(* IEC 61131-3 sources: NachHouse_TST/API/pilot_Api_V11 (part 2) *)

(* ---- 03_Nh_Api_ENGINE.st ---- *)
// Single-owner transaction engine, snapshots, diffs and room operations.
// SK: Transakcny automat jedneho vlastnika, snapshoty, diffy a room operacie.

FUNCTION NhApiClearRoom : BOOL
   // Clears configuration and state of one internal room slot. SK: Vynuluje konfiguraciu a stav jedneho interneho room slotu.
   VAR_INPUT
      Index : UINT; // Internal model-device slot 1..800. SK: Interny slot modeloveho zariadenia 1..800.
   END_VAR
   NhRoomsConfig[Index].Used := FALSE;
   NhRoomsConfig[Index].RoomId := 0;
   NhRoomsConfig[Index].Name := '';
   NhRoomsConfig[Index].ProjectName := '';
   NhRoomsConfig[Index].IconId := 0;
   NhRoomsConfig[Index].SortDefault := 0;
   NhRoomsState[Index].RoomId := 0;
   NhRoomsState[Index].Temperature := 0.0;
   NhRoomsState[Index].Humidity := 0.0;
   NhRoomsState[Index].Presence := FALSE;
   NhRoomsState[Index].DayPhase := 140;
   NhRoomsState[Index].CategoryMask := 0;
   NhRoomsState[Index].AlarmLevel := 0;
   NhRoomsState[Index].Online := FALSE;
   NhRoomsState[Index].Twilight := FALSE;
   NhApiClearRoom := TRUE;
END_FUNCTION

FUNCTION NhApiInitialize : BOOL
   // Initializes API buffers, handshake and deterministic pilot data once. SK: Jednorazovo inicializuje API buffery, handshake a deterministicke pilotne data.
   VAR
      Index : UINT; // Initialization index. SK: Inicializacny index.
   END_VAR
   NhApiInitialize := NhApiInitialized;
   IF NhApiInitialized THEN RETURN; END_IF;

   NhApiClearBuffer(Buffer := ADR(NhApiTX), Length := NH_API_TX_BYTE_CAPACITY);
   NhApiClearBuffer(Buffer := ADR(NhApiRX), Length := NH_API_RX_BYTE_CAPACITY);
   FOR Index := 1 TO NH_API_MAX_ROOMS DO
      NhApiClearRoom(Index := Index);
   END_FOR;

   FOR Index := 1 TO 30 DO
      NhRoomsConfig[Index].Used := TRUE;
      NhRoomsConfig[Index].RoomId := UINT_TO_UDINT(Index);
      NhRoomsConfig[Index].ProjectName := 'TEST';
      NhRoomsConfig[Index].IconId := SEL(Index >= 26, 16, 19);
      NhRoomsConfig[Index].SortDefault := Index;
      CASE Index OF
         1: NhRoomsConfig[Index].Name := 'Hall 1'; NhRoomsConfig[Index].ProjectName := '1.08';
         2: NhRoomsConfig[Index].Name := 'Kitchen'; NhRoomsConfig[Index].ProjectName := '1.07';
         3: NhRoomsConfig[Index].Name := 'Corridor 1'; NhRoomsConfig[Index].ProjectName := '1.04';
         4: NhRoomsConfig[Index].Name := 'Bathroom 1'; NhRoomsConfig[Index].ProjectName := '1.06';
         5: NhRoomsConfig[Index].Name := 'WC'; NhRoomsConfig[Index].ProjectName := '1.05';
         6: NhRoomsConfig[Index].Name := 'Bedroom'; NhRoomsConfig[Index].ProjectName := '1.09';
         7: NhRoomsConfig[Index].Name := 'Boiler'; NhRoomsConfig[Index].ProjectName := '1.03';
         8: NhRoomsConfig[Index].Name := 'Living room'; NhRoomsConfig[Index].ProjectName := '1.01';
         9: NhRoomsConfig[Index].Name := 'Corridor 1F'; NhRoomsConfig[Index].ProjectName := '1.02';
         10: NhRoomsConfig[Index].Name := 'Room 2.07'; NhRoomsConfig[Index].ProjectName := '2.07';
         11: NhRoomsConfig[Index].Name := 'Kitchen 2F'; NhRoomsConfig[Index].ProjectName := '2.03';
         12: NhRoomsConfig[Index].Name := 'Room 2.06'; NhRoomsConfig[Index].ProjectName := '2.06';
         13: NhRoomsConfig[Index].Name := 'Bathroom 2F'; NhRoomsConfig[Index].ProjectName := '2.05';
         14: NhRoomsConfig[Index].Name := 'Entrance hall'; NhRoomsConfig[Index].ProjectName := '0.01';
         15: NhRoomsConfig[Index].Name := 'Garage'; NhRoomsConfig[Index].ProjectName := '0.02';
         16: NhRoomsConfig[Index].Name := 'Storage'; NhRoomsConfig[Index].ProjectName := '0.03';
         17: NhRoomsConfig[Index].Name := 'Basement corridor'; NhRoomsConfig[Index].ProjectName := '0.04';
         18: NhRoomsConfig[Index].Name := 'Office'; NhRoomsConfig[Index].ProjectName := '1.10';
         19: NhRoomsConfig[Index].Name := 'Wardrobe'; NhRoomsConfig[Index].ProjectName := '1.11';
         20: NhRoomsConfig[Index].Name := 'Fitness'; NhRoomsConfig[Index].ProjectName := '0.06';
         21: NhRoomsConfig[Index].Name := 'Technical'; NhRoomsConfig[Index].ProjectName := '0.07';
         22: NhRoomsConfig[Index].Name := 'Wine room'; NhRoomsConfig[Index].ProjectName := '0.08';
         23: NhRoomsConfig[Index].Name := 'Guest room'; NhRoomsConfig[Index].ProjectName := '2.01';
         24: NhRoomsConfig[Index].Name := 'Children 1'; NhRoomsConfig[Index].ProjectName := '2.02';
         25: NhRoomsConfig[Index].Name := 'Children 2'; NhRoomsConfig[Index].ProjectName := '2.04';
         26: NhRoomsConfig[Index].Name := 'Terrace'; NhRoomsConfig[Index].ProjectName := 'E.01';
         27: NhRoomsConfig[Index].Name := 'Gazebo'; NhRoomsConfig[Index].ProjectName := 'E.02';
         28: NhRoomsConfig[Index].Name := 'Pool'; NhRoomsConfig[Index].ProjectName := 'E.03';
         29: NhRoomsConfig[Index].Name := 'Garden'; NhRoomsConfig[Index].ProjectName := 'E.04';
         30: NhRoomsConfig[Index].Name := 'Sauna'; NhRoomsConfig[Index].ProjectName := '0.09';
      END_CASE;
      NhRoomsState[Index].RoomId := UINT_TO_UDINT(Index);
      NhRoomsState[Index].Temperature := 20.0 + UINT_TO_REAL(Index) * 0.1;
      NhRoomsState[Index].Humidity := 40.0 + UINT_TO_REAL(Index MOD 15);
      NhRoomsState[Index].Presence := (Index MOD 4) = 0;
      CASE Index MOD 4 OF
         0: NhRoomsState[Index].DayPhase := 140;
         1: NhRoomsState[Index].DayPhase := 142;
         2: NhRoomsState[Index].DayPhase := 144;
         3: NhRoomsState[Index].DayPhase := 146;
      END_CASE;
      NhRoomsState[Index].CategoryMask := UINT_TO_DWORD(Index MOD 8);
      NhRoomsState[Index].AlarmLevel := 0;
      NhRoomsState[Index].Online := (Index MOD 3) <> 0;
      NhRoomsState[Index].Twilight := (Index MOD 3) <> 1;
   END_FOR;

   FOR Index := 1 TO NH_API_MAX_ROOMS DO
      NhConfigShadow[Index] := NhRoomsConfig[Index];
      NhStateShadow[Index] := NhRoomsState[Index];
   END_FOR;

   // Deterministic compact LOAD_800 device model. SK: Deterministicky kompaktny model 800 zariadeni.
   FOR Index := 1 TO NH_LOAD_DEVICE_COUNT DO
      IF Index <= 300 THEN
         NhLoadDevices[Index] := 16#01000064; // light, level 100
      ELSIF Index <= 420 THEN
         NhLoadDevices[Index] := 16#02000064; // roller, position 100
      ELSIF Index <= 520 THEN
         NhLoadDevices[Index] := 16#030000D2; // heating, 21.0 C
      ELSIF Index <= 600 THEN
         NhLoadDevices[Index] := 16#040000DC; // climate, 22.0 C
      ELSIF Index <= 640 THEN
         NhLoadDevices[Index] := 16#05000001; // water, enabled
      ELSE
         NhLoadDevices[Index] := 16#06000000 OR UINT_TO_DWORD(Index MOD 256); // sensor control group
      END_IF;
   END_FOR;

   NhApiInfo.ApiVersion := NH_API_VERSION;
   NhApiInfo.OwnerClientId := 0;
   NhApiInfo.State := NH_API_STATE_IDLE;
   NhActiveOwnerClientId := 0;
   NhExpectedState := NH_API_STATE_IDLE;
   NhTransactionMode := NH_API_MODE_NONE;
   NhTransactionLastMs := NhApiSystemTimeMs();
   NhPublishedFrameId := 0;
   NhCommandResult := NH_API_RESULT_NONE;
   NhResultPending := FALSE;
   NhPendingConfigCount := 0;
   NhPendingStateCount := 0;
   NhSnapshotActive := FALSE;

   NhApiTest.Execute := FALSE;
   NhApiTest.Finished := FALSE;
   NhApiTest.Action := NH_API_TEST_NONE;
   NhApiTest.ResultCode := NH_API_RESULT_NONE;
   NhLoadTest.DepartureActive := FALSE;
   NhLoadTest.LastChangedCount := 0;
   NhLoadTest.LastApplyMs := 0;
   NhLoadTest.Sequence := 0;
   NhApiInitialized := TRUE;
   NhApiInitialize := TRUE;
END_FUNCTION

FUNCTION NhApiBeginFrame : BOOL
   // Clears TX and writes the fixed 40-byte frame header. SK: Vycisti TX a zapise pevnu 40-bajtovu hlavicku ramca.
   VAR_INPUT
      MessageType  : UINT;  // NH_API_MSG_* value. SK: Hodnota NH_API_MSG_*.
      SchemaId     : UINT;  // NH_API_SCHEMA_* value. SK: Hodnota NH_API_SCHEMA_*.
      OwnerClientId: UDINT; // Target owner token; zero is broadcast. SK: Cielovy token vlastnika; nula je broadcast.
      RecordCount  : UINT;  // Number of payload records. SK: Pocet zaznamov payloadu.
      RecordSize   : UINT;  // Fixed size of one payload record. SK: Pevna velkost jedneho payload zaznamu.
      PartIndex    : UINT;  // One-based part index. SK: Index casti cislovany od jedna.
      PartCount    : UINT;  // Total parts in this section. SK: Celkovy pocet casti sekcie.
      ResultCode   : USINT; // NH_API_RESULT_* value. SK: Hodnota NH_API_RESULT_*.
   END_VAR
   VAR
      Buffer      : PTR_TO BYTE; // Byte view of NhApiTX. SK: Bajtovy pohlad na NhApiTX.
      PayloadSize : UDINT;       // Calculated payload size. SK: Vypocitana velkost payloadu.
      TotalSize   : UDINT;       // Header plus payload size. SK: Velkost hlavicky a payloadu.
   END_VAR
   Buffer := ADR(NhApiTX);
   NhApiClearBuffer(Buffer := Buffer, Length := NH_API_TX_BYTE_CAPACITY);
   PayloadSize := UINT_TO_UDINT(RecordCount) * UINT_TO_UDINT(RecordSize);
   TotalSize := UINT_TO_UDINT(NH_API_HEADER_SIZE) + PayloadSize;
   IF TotalSize > UINT_TO_UDINT(NH_API_TX_BYTE_CAPACITY) THEN
      NhApiBeginFrame := FALSE;
      RETURN;
   END_IF;
   NhApiWriteU32(Buffer := Buffer, Offset := 0, Value := DWORD_TO_UDINT(NH_API_MAGIC));
   NhApiWriteU16(Buffer := Buffer, Offset := 4, Value := NH_API_VERSION);
   NhApiWriteU16(Buffer := Buffer, Offset := 6, Value := NH_API_HEADER_SIZE);
   NhApiWriteU16(Buffer := Buffer, Offset := 8, Value := MessageType);
   NhApiWriteU16(Buffer := Buffer, Offset := 10, Value := SchemaId);
   NhApiWriteU32(Buffer := Buffer, Offset := 12, Value := OwnerClientId);
   NhApiWriteU16(Buffer := Buffer, Offset := 16, Value := RecordCount);
   NhApiWriteU16(Buffer := Buffer, Offset := 18, Value := RecordSize);
   NhApiWriteByte(Buffer := Buffer, Offset := 20, Value := WORD_TO_BYTE(UINT_TO_WORD(PartIndex)));
   NhApiWriteByte(Buffer := Buffer, Offset := 21, Value := WORD_TO_BYTE(UINT_TO_WORD(PartCount)));
   NhApiWriteByte(Buffer := Buffer, Offset := 22, Value := USINT_TO_BYTE(ResultCode));
   NhApiWriteByte(Buffer := Buffer, Offset := 23, Value := 0);
   NhApiWriteU32(Buffer := Buffer, Offset := 24, Value := PayloadSize);
   NhApiWriteU32(Buffer := Buffer, Offset := 28, Value := TotalSize);
   NhApiWriteU32(Buffer := Buffer, Offset := 32, Value := 0);
   NhApiWriteU32(Buffer := Buffer, Offset := 36, Value := 0);
   NhApiBeginFrame := TRUE;
END_FUNCTION

FUNCTION NhApiPublishFrame : BOOL
   // Adds CRC and publishes TX by changing State only after the buffer is stable. SK: Doplni CRC a publikuje TX zmenou State az po ustaleni buffera.
   VAR_INPUT
      NextState : UINT; // New persistent handshake step. SK: Novy trvaly handshake krok.
   END_VAR
   VAR
      Buffer    : PTR_TO BYTE; // Byte view of NhApiTX. SK: Bajtovy pohlad na NhApiTX.
      TotalSize : UINT;        // Valid frame byte count. SK: Pocet platnych bajtov ramca.
      Crc       : DWORD;       // CRC32 of the frame. SK: CRC32 ramca.
   END_VAR
   Buffer := ADR(NhApiTX);
   TotalSize := UDINT_TO_UINT(NhApiReadU32(Buffer := Buffer, Offset := 28));
   NhPublishedFrameId := NhPublishedFrameId + 1;
   IF NhPublishedFrameId = 0 THEN NhPublishedFrameId := 1; END_IF;
   NhApiWriteU32(Buffer := Buffer, Offset := 32, Value := NhPublishedFrameId);
   Crc := NhApiFrameCrc32(Buffer := Buffer, Length := TotalSize);
   NhApiWriteU32(Buffer := Buffer, Offset := 36, Value := DWORD_TO_UDINT(Crc));
   NhExpectedState := NextState;
   NhTransactionLastMs := NhApiSystemTimeMs();
   NhApiInfo.State := NextState;
   NhApiPublishFrame := TRUE;
END_FUNCTION

FUNCTION NhApiResetTransaction : BOOL
   // Releases the global mailbox and clears internal sequence state. SK: Uvolni globalny mailbox a vycisti interny stav sekvencie.
   NhApiInfo.OwnerClientId := 0;
   NhApiInfo.State := NH_API_STATE_IDLE;
   NhActiveOwnerClientId := 0;
   NhExpectedState := NH_API_STATE_IDLE;
   NhTransactionMode := NH_API_MODE_NONE;
   NhTransactionLastMs := NhApiSystemTimeMs();
   NhCommandResult := NH_API_RESULT_NONE;
   NhResultPending := FALSE;
   NhPendingConfigCount := 0;
   NhPendingStateCount := 0;
   NhSnapshotActive := FALSE;
   NhApiResetTransaction := TRUE;
END_FUNCTION

FUNCTION NhApiApplyAdd : USINT
   // Adds a room to the first free internal slot. SK: Prida miestnost do prveho volneho interneho slotu.
   VAR_INPUT
      Record : NH_ROOM_CONFIG; // New room configuration. SK: Konfiguracia novej miestnosti.
   END_VAR
   VAR
      Slot : UINT; // Free internal room slot. SK: Volny interny room slot.
   END_VAR
   IF (Record.RoomId = 0) OR (LEN(Record.Name) = 0) THEN NhApiApplyAdd := NH_API_RESULT_INVALID; RETURN; END_IF;
   IF NhApiFindRoom(RoomId := Record.RoomId) <> 0 THEN NhApiApplyAdd := NH_API_RESULT_ALREADY_EXISTS; RETURN; END_IF;
   Slot := NhApiFindFreeRoom();
   IF Slot = 0 THEN NhApiApplyAdd := NH_API_RESULT_NO_FREE_SLOT; RETURN; END_IF;
   NhRoomsConfig[Slot] := Record;
   NhRoomsConfig[Slot].Used := TRUE;
   IF NhRoomsConfig[Slot].IconId = 0 THEN NhRoomsConfig[Slot].IconId := 16; END_IF;
   IF NhRoomsConfig[Slot].SortDefault = 0 THEN NhRoomsConfig[Slot].SortDefault := Slot; END_IF;
   NhRoomsState[Slot].RoomId := Record.RoomId;
   NhRoomsState[Slot].Temperature := 20.0;
   NhRoomsState[Slot].Humidity := 40.0;
   NhRoomsState[Slot].Presence := FALSE;
   NhRoomsState[Slot].DayPhase := 140;
   NhRoomsState[Slot].CategoryMask := 0;
   NhRoomsState[Slot].AlarmLevel := 0;
   NhRoomsState[Slot].Online := TRUE;
   NhRoomsState[Slot].Twilight := FALSE;
   NhApiApplyAdd := NH_API_RESULT_OK;
END_FUNCTION

FUNCTION NhApiApplyDelete : USINT
   // Deletes a room by stable RoomId. SK: Zmaze miestnost podla stabilneho RoomId.
   VAR_INPUT
      RoomId : UDINT; // ID of the room to delete. SK: ID mazanej miestnosti.
   END_VAR
   VAR
      Slot : UINT;   // Located internal slot. SK: Najdeny interny slot.
   END_VAR
   Slot := NhApiFindRoom(RoomId := RoomId);
   IF Slot = 0 THEN NhApiApplyDelete := NH_API_RESULT_NOT_FOUND; RETURN; END_IF;
   NhApiClearRoom(Index := Slot);
   NhApiApplyDelete := NH_API_RESULT_OK;
END_FUNCTION

FUNCTION NhApiApplyConfig : USINT
   // Replaces complete configuration of an existing room. SK: Nahradi celu konfiguraciu existujucej miestnosti.
   VAR_INPUT
      Record : NH_ROOM_CONFIG; // Complete new configuration. SK: Uplna nova konfiguracia.
   END_VAR
   VAR
      Slot : UINT;            // Located internal slot. SK: Najdeny interny slot.
   END_VAR
   Slot := NhApiFindRoom(RoomId := Record.RoomId);
   IF Slot = 0 THEN NhApiApplyConfig := NH_API_RESULT_NOT_FOUND; RETURN; END_IF;
   IF LEN(Record.Name) = 0 THEN NhApiApplyConfig := NH_API_RESULT_INVALID; RETURN; END_IF;
   NhRoomsConfig[Slot] := Record;
   NhRoomsConfig[Slot].Used := TRUE;
   NhApiApplyConfig := NH_API_RESULT_OK;
END_FUNCTION

FUNCTION NhApiApplyState : USINT
   // Replaces complete dynamic state of an existing room. SK: Nahradi cely dynamicky stav existujucej miestnosti.
   VAR_INPUT
      Record : NH_ROOM_STATE; // Complete new state. SK: Uplny novy stav.
   END_VAR
   VAR
      Slot : UINT;           // Located internal slot. SK: Najdeny interny slot.
   END_VAR
   Slot := NhApiFindRoom(RoomId := Record.RoomId);
   IF Slot = 0 THEN NhApiApplyState := NH_API_RESULT_NOT_FOUND; RETURN; END_IF;
   IF (Record.Temperature < -50.0) OR (Record.Temperature > 100.0) OR
      (Record.Humidity < 0.0) OR (Record.Humidity > 100.0) OR (Record.AlarmLevel > 2) THEN
      NhApiApplyState := NH_API_RESULT_INVALID;
      RETURN;
   END_IF;
   NhRoomsState[Slot] := Record;
   NhApiApplyState := NH_API_RESULT_OK;
END_FUNCTION

FUNCTION NhApiApplyCopy : USINT
   // Copies an existing room into a new RoomId. SK: Skopiruje existujucu miestnost do noveho RoomId.
   VAR_INPUT
      SourceRoomId : UDINT;         // Source room ID. SK: ID zdrojovej miestnosti.
      Target       : NH_ROOM_CONFIG;// Target ID and optional replacements. SK: Cielove ID a volitelne nahrady.
   END_VAR
   VAR
      SourceSlot : UINT; // Source internal slot. SK: Zdrojovy interny slot.
      TargetSlot : UINT; // Target free slot. SK: Cielovy volny slot.
   END_VAR
   SourceSlot := NhApiFindRoom(RoomId := SourceRoomId);
   IF SourceSlot = 0 THEN NhApiApplyCopy := NH_API_RESULT_NOT_FOUND; RETURN; END_IF;
   IF Target.RoomId = 0 THEN NhApiApplyCopy := NH_API_RESULT_INVALID; RETURN; END_IF;
   IF NhApiFindRoom(RoomId := Target.RoomId) <> 0 THEN NhApiApplyCopy := NH_API_RESULT_ALREADY_EXISTS; RETURN; END_IF;
   TargetSlot := NhApiFindFreeRoom();
   IF TargetSlot = 0 THEN NhApiApplyCopy := NH_API_RESULT_NO_FREE_SLOT; RETURN; END_IF;
   NhRoomsConfig[TargetSlot] := NhRoomsConfig[SourceSlot];
   NhRoomsConfig[TargetSlot].RoomId := Target.RoomId;
   NhRoomsConfig[TargetSlot].SortDefault := TargetSlot;
   IF LEN(Target.Name) > 0 THEN NhRoomsConfig[TargetSlot].Name := Target.Name; END_IF;
   IF LEN(Target.ProjectName) > 0 THEN NhRoomsConfig[TargetSlot].ProjectName := Target.ProjectName; END_IF;
   IF Target.IconId > 0 THEN NhRoomsConfig[TargetSlot].IconId := Target.IconId; END_IF;
   NhRoomsState[TargetSlot] := NhRoomsState[SourceSlot];
   NhRoomsState[TargetSlot].RoomId := Target.RoomId;
   NhApiApplyCopy := NH_API_RESULT_OK;
END_FUNCTION

FUNCTION NhApiCaptureConfigChanges : BOOL
   // Freezes all unpublished configuration changes. SK: Zmrazi vsetky nepublikovane zmeny konfiguracie.
   VAR
      Index : UINT; // Scanned room slot. SK: Prehladavany room slot.
   END_VAR
   NhPendingConfigCount := 0;
   FOR Index := 1 TO NH_API_MAX_ROOMS DO
      IF NOT NhApiConfigEqual(A := NhRoomsConfig[Index], B := NhConfigShadow[Index]) THEN
         NhPendingConfigCount := NhPendingConfigCount + 1;
         IF NhRoomsConfig[Index].Used THEN
            NhPendingConfigOperation[NhPendingConfigCount] := NH_API_CHANGE_UPSERT;
            NhPendingConfigRoomId[NhPendingConfigCount] := NhRoomsConfig[Index].RoomId;
         ELSE
            NhPendingConfigOperation[NhPendingConfigCount] := NH_API_CHANGE_DELETE;
            NhPendingConfigRoomId[NhPendingConfigCount] := NhConfigShadow[Index].RoomId;
         END_IF;
         NhPendingConfig[NhPendingConfigCount] := NhRoomsConfig[Index];
         NhConfigShadow[Index] := NhRoomsConfig[Index];
      END_IF;
   END_FOR;
   NhPendingConfigNext := 1;
   NhPendingConfigPart := 1;
   NhPendingConfigParts := 0;
   IF NhPendingConfigCount > 0 THEN
      NhPendingConfigParts := (NhPendingConfigCount + NH_API_CONFIG_DIFF_PER_FRAME - 1) / NH_API_CONFIG_DIFF_PER_FRAME;
   END_IF;
   NhApiCaptureConfigChanges := NhPendingConfigCount > 0;
END_FUNCTION

FUNCTION NhApiCaptureStateChanges : BOOL
   // Freezes all unpublished dynamic-state changes. SK: Zmrazi vsetky nepublikovane zmeny dynamickeho stavu.
   VAR
      Index : UINT; // Scanned room slot. SK: Prehladavany room slot.
   END_VAR
   NhPendingStateCount := 0;
   FOR Index := 1 TO NH_API_MAX_ROOMS DO
      IF NOT NhApiStateEqual(A := NhRoomsState[Index], B := NhStateShadow[Index]) THEN
         NhPendingStateCount := NhPendingStateCount + 1;
         IF NhRoomsConfig[Index].Used THEN
            NhPendingStateOperation[NhPendingStateCount] := NH_API_CHANGE_UPSERT;
            NhPendingStateRoomId[NhPendingStateCount] := NhRoomsState[Index].RoomId;
         ELSE
            NhPendingStateOperation[NhPendingStateCount] := NH_API_CHANGE_DELETE;
            NhPendingStateRoomId[NhPendingStateCount] := NhStateShadow[Index].RoomId;
         END_IF;
         NhPendingState[NhPendingStateCount] := NhRoomsState[Index];
         NhStateShadow[Index] := NhRoomsState[Index];
      END_IF;
   END_FOR;
   NhPendingStateNext := 1;
   NhPendingStatePart := 1;
   NhPendingStateParts := 0;
   IF NhPendingStateCount > 0 THEN
      NhPendingStateParts := (NhPendingStateCount + NH_API_STATE_DIFF_PER_FRAME - 1) / NH_API_STATE_DIFF_PER_FRAME;
   END_IF;
   NhApiCaptureStateChanges := NhPendingStateCount > 0;
END_FUNCTION

FUNCTION NhApiCaptureAllChanges : BOOL
   // Freezes current config and state changes in one PLC cycle. SK: Zmrazi aktualne config a state zmeny v jednom PLC cykle.
   VAR
      ConfigChanged : BOOL; // At least one config changed. SK: Zmenil sa aspon jeden config.
      StateChanged  : BOOL; // At least one state changed. SK: Zmenil sa aspon jeden state.
   END_VAR
   ConfigChanged := NhApiCaptureConfigChanges();
   StateChanged := NhApiCaptureStateChanges();
   NhApiCaptureAllChanges := ConfigChanged OR StateChanged;
END_FUNCTION

FUNCTION NhApiStartSnapshot : BOOL
   // Freezes the authoritative room image for a complete snapshot. SK: Zmrazi autoritativny obraz miestnosti pre kompletny snapshot.
   VAR
      Index : UINT; // Scanned source room slot. SK: Prehladavany zdrojovy room slot.
   END_VAR
   NhSnapshotCount := 0;
   FOR Index := 1 TO NH_API_MAX_ROOMS DO
      IF NhRoomsConfig[Index].Used THEN
         NhSnapshotCount := NhSnapshotCount + 1;
         NhSnapshotConfig[NhSnapshotCount] := NhRoomsConfig[Index];
         NhSnapshotState[NhSnapshotCount] := NhRoomsState[Index];
      END_IF;
      // The frozen snapshot is the new cache baseline; later PLC changes become diffs. SK: Zmrazeny snapshot je novy zaklad cache; neskorsie PLC zmeny sa stanu diffom.
      NhConfigShadow[Index] := NhRoomsConfig[Index];
      NhStateShadow[Index] := NhRoomsState[Index];
   END_FOR;
   NhPendingConfigCount := 0;
   NhPendingStateCount := 0;
   NhSnapshotActive := TRUE;
   NhSnapshotStage := 1;
   NhSnapshotNext := 1;
   NhSnapshotPart := 1;
   NhSnapshotParts := (NhSnapshotCount + NH_API_CONFIG_PER_FRAME - 1) / NH_API_CONFIG_PER_FRAME;
   IF NhSnapshotParts = 0 THEN NhSnapshotParts := 1; END_IF;
   NhApiStartSnapshot := TRUE;
END_FUNCTION

FUNCTION NhApiBuildNextSnapshotFrame : BOOL
   // Builds the next CONFIG, STATE or DONE snapshot frame without publishing State yet. SK: Vytvori dalsi CONFIG, STATE alebo DONE snapshot ramec bez publikovania State.
   VAR
      Buffer : PTR_TO BYTE; // Byte view of NhApiTX. SK: Bajtovy pohlad na NhApiTX.
      Count  : USINT;       // Records in this frame. SK: Pocet zaznamov v tomto ramci.
      Index  : USINT;       // Local record index. SK: Lokalny index zaznamu.
      Source : USINT;       // Frozen snapshot index. SK: Index zmrazeneho snapshotu.
      Offset : UINT;        // Record byte offset. SK: Bajtovy offset zaznamu.
   END_VAR
   NhApiBuildNextSnapshotFrame := FALSE;
   IF NOT NhSnapshotActive THEN RETURN; END_IF;
   Buffer := ADR(NhApiTX);

   IF NhSnapshotStage = 1 THEN
      Count := NH_API_CONFIG_PER_FRAME;
      IF NhSnapshotCount = 0 THEN
         Count := 0;
      ELSIF (NhSnapshotNext + Count - 1) > NhSnapshotCount THEN
         Count := NhSnapshotCount - NhSnapshotNext + 1;
      END_IF;
      NhApiBeginFrame(MessageType := NH_API_MSG_CONFIG_SNAPSHOT, SchemaId := NH_API_SCHEMA_ROOM_CONFIG,
         OwnerClientId := NhActiveOwnerClientId, RecordCount := USINT_TO_UINT(Count),
         RecordSize := NH_API_CONFIG_RECORD_SIZE, PartIndex := USINT_TO_UINT(NhSnapshotPart),
         PartCount := USINT_TO_UINT(NhSnapshotParts), ResultCode := NH_API_RESULT_OK);
      IF Count > 0 THEN
         FOR Index := 0 TO Count - 1 DO
            Source := NhSnapshotNext + Index;
            Offset := NH_API_HEADER_SIZE + USINT_TO_UINT(Index) * NH_API_CONFIG_RECORD_SIZE;
            NhApiWriteConfigRecord(Buffer := Buffer, Offset := Offset, Record := NhSnapshotConfig[Source]);
         END_FOR;
      END_IF;
      NhSnapshotNext := NhSnapshotNext + Count;
      NhSnapshotPart := NhSnapshotPart + 1;
      IF (NhSnapshotCount = 0) OR (NhSnapshotNext > NhSnapshotCount) THEN
         NhSnapshotStage := 2;
         NhSnapshotNext := 1;
         NhSnapshotPart := 1;
         NhSnapshotParts := (NhSnapshotCount + NH_API_STATE_PER_FRAME - 1) / NH_API_STATE_PER_FRAME;
         IF NhSnapshotParts = 0 THEN NhSnapshotParts := 1; END_IF;
      END_IF;
      NhApiBuildNextSnapshotFrame := TRUE;
      RETURN;
   END_IF;

   IF NhSnapshotStage = 2 THEN
      Count := NH_API_STATE_PER_FRAME;
      IF NhSnapshotCount = 0 THEN
         Count := 0;
      ELSIF (NhSnapshotNext + Count - 1) > NhSnapshotCount THEN
         Count := NhSnapshotCount - NhSnapshotNext + 1;
      END_IF;
      NhApiBeginFrame(MessageType := NH_API_MSG_STATE_SNAPSHOT, SchemaId := NH_API_SCHEMA_ROOM_STATE,
         OwnerClientId := NhActiveOwnerClientId, RecordCount := USINT_TO_UINT(Count),
         RecordSize := NH_API_STATE_RECORD_SIZE, PartIndex := USINT_TO_UINT(NhSnapshotPart),
         PartCount := USINT_TO_UINT(NhSnapshotParts), ResultCode := NH_API_RESULT_OK);
      IF Count > 0 THEN
         FOR Index := 0 TO Count - 1 DO
            Source := NhSnapshotNext + Index;
            Offset := NH_API_HEADER_SIZE + USINT_TO_UINT(Index) * NH_API_STATE_RECORD_SIZE;
            NhApiWriteStateRecord(Buffer := Buffer, Offset := Offset, Record := NhSnapshotState[Source]);
         END_FOR;
      END_IF;
      NhSnapshotNext := NhSnapshotNext + Count;
      NhSnapshotPart := NhSnapshotPart + 1;
      IF (NhSnapshotCount = 0) OR (NhSnapshotNext > NhSnapshotCount) THEN
         NhSnapshotStage := 3;
      END_IF;
      NhApiBuildNextSnapshotFrame := TRUE;
      RETURN;
   END_IF;

   IF NhSnapshotStage = 3 THEN
      NhApiBeginFrame(MessageType := NH_API_MSG_SNAPSHOT_DONE, SchemaId := NH_API_SCHEMA_NONE,
         OwnerClientId := NhActiveOwnerClientId, RecordCount := 0, RecordSize := 0,
         PartIndex := 1, PartCount := 1, ResultCode := NH_API_RESULT_OK);
      NhSnapshotStage := 4;
      NhApiBuildNextSnapshotFrame := TRUE;
      RETURN;
   END_IF;

   NhSnapshotActive := FALSE;
END_FUNCTION

FUNCTION NhApiBuildNextDiffFrame : BOOL
   // Builds the next frozen CONFIG or STATE diff frame. SK: Vytvori dalsi zmrazeny CONFIG alebo STATE diff ramec.
   VAR
      Buffer : PTR_TO BYTE; // Byte view of NhApiTX. SK: Bajtovy pohlad na NhApiTX.
      Count  : USINT;       // Changes in this frame. SK: Pocet zmien v tomto ramci.
      Index  : USINT;       // Local change index. SK: Lokalny index zmeny.
      Source : USINT;       // Frozen change index. SK: Index zmrazenej zmeny.
      Offset : UINT;        // Change byte offset. SK: Bajtovy offset zmeny.
   END_VAR
   NhApiBuildNextDiffFrame := FALSE;
   Buffer := ADR(NhApiTX);

   IF NhPendingConfigNext <= NhPendingConfigCount THEN
      Count := NH_API_CONFIG_DIFF_PER_FRAME;
      IF (NhPendingConfigNext + Count - 1) > NhPendingConfigCount THEN
         Count := NhPendingConfigCount - NhPendingConfigNext + 1;
      END_IF;
      NhApiBeginFrame(MessageType := NH_API_MSG_CONFIG_DIFF, SchemaId := NH_API_SCHEMA_ROOM_CONFIG,
         OwnerClientId := NhActiveOwnerClientId, RecordCount := USINT_TO_UINT(Count),
         RecordSize := NH_API_CONFIG_DIFF_SIZE, PartIndex := USINT_TO_UINT(NhPendingConfigPart),
         PartCount := USINT_TO_UINT(NhPendingConfigParts), ResultCode := NhCommandResult);
      FOR Index := 0 TO Count - 1 DO
         Source := NhPendingConfigNext + Index;
         Offset := NH_API_HEADER_SIZE + USINT_TO_UINT(Index) * NH_API_CONFIG_DIFF_SIZE;
         NhApiWriteByte(Buffer := Buffer, Offset := Offset, Value := USINT_TO_BYTE(NhPendingConfigOperation[Source]));
         NhApiWriteU32(Buffer := Buffer, Offset := Offset + 1, Value := NhPendingConfigRoomId[Source]);
         NhApiWriteConfigRecord(Buffer := Buffer, Offset := Offset + 5, Record := NhPendingConfig[Source]);
      END_FOR;
      NhPendingConfigNext := NhPendingConfigNext + Count;
      NhPendingConfigPart := NhPendingConfigPart + 1;
      NhApiBuildNextDiffFrame := TRUE;
      RETURN;
   END_IF;

   IF NhPendingStateNext <= NhPendingStateCount THEN
      Count := NH_API_STATE_DIFF_PER_FRAME;
      IF (NhPendingStateNext + Count - 1) > NhPendingStateCount THEN
         Count := NhPendingStateCount - NhPendingStateNext + 1;
      END_IF;
      NhApiBeginFrame(MessageType := NH_API_MSG_STATE_DIFF, SchemaId := NH_API_SCHEMA_ROOM_STATE,
         OwnerClientId := NhActiveOwnerClientId, RecordCount := USINT_TO_UINT(Count),
         RecordSize := NH_API_STATE_DIFF_SIZE, PartIndex := USINT_TO_UINT(NhPendingStatePart),
         PartCount := USINT_TO_UINT(NhPendingStateParts), ResultCode := NhCommandResult);
      FOR Index := 0 TO Count - 1 DO
         Source := NhPendingStateNext + Index;
         Offset := NH_API_HEADER_SIZE + USINT_TO_UINT(Index) * NH_API_STATE_DIFF_SIZE;
         NhApiWriteByte(Buffer := Buffer, Offset := Offset, Value := USINT_TO_BYTE(NhPendingStateOperation[Source]));
         NhApiWriteU32(Buffer := Buffer, Offset := Offset + 1, Value := NhPendingStateRoomId[Source]);
         NhApiWriteStateRecord(Buffer := Buffer, Offset := Offset + 5, Record := NhPendingState[Source]);
      END_FOR;
      NhPendingStateNext := NhPendingStateNext + Count;
      NhPendingStatePart := NhPendingStatePart + 1;
      NhApiBuildNextDiffFrame := TRUE;
      RETURN;
   END_IF;
END_FUNCTION

FUNCTION NhApiBuildResultFrame : BOOL
   // Builds the final command result frame. SK: Vytvori posledny ramec vysledku prikazu.
   NhApiBuildResultFrame := FALSE;
   IF NOT NhResultPending THEN RETURN; END_IF;
   NhApiBeginFrame(MessageType := NH_API_MSG_RESULT, SchemaId := NH_API_SCHEMA_NONE,
      OwnerClientId := NhActiveOwnerClientId, RecordCount := 0, RecordSize := 0,
      PartIndex := 1, PartCount := 1, ResultCode := NhCommandResult);
   NhResultPending := FALSE;
   NhApiBuildResultFrame := TRUE;
END_FUNCTION

FUNCTION NhApiBuildNextFrame : BOOL
   // Selects and builds the next frame of the active sequence. SK: Vyberie a vytvori dalsi ramec aktivnej sekvencie.
   NhApiBuildNextFrame := FALSE;
   IF (NhTransactionMode = NH_API_MODE_SNAPSHOT) OR (NhTransactionMode = NH_API_MODE_BROADCAST_SNAPSHOT) THEN
      NhApiBuildNextFrame := NhApiBuildNextSnapshotFrame();
      RETURN;
   END_IF;
   IF (NhTransactionMode = NH_API_MODE_COMMAND) OR (NhTransactionMode = NH_API_MODE_BROADCAST_DIFF) THEN
      IF NhApiBuildNextDiffFrame() THEN
         NhApiBuildNextFrame := TRUE;
         RETURN;
      END_IF;
      IF NhTransactionMode = NH_API_MODE_COMMAND THEN
         NhApiBuildNextFrame := NhApiBuildResultFrame();
      END_IF;
   END_IF;
END_FUNCTION

FUNCTION NhApiPublishNextTargetFrame : BOOL
   // Publishes the next targeted frame or releases the transaction after the final ACK. SK: Publikuje dalsi cielovy ramec alebo po poslednom ACK uvolni transakciu.
   VAR
      NextState : UINT; // Next odd PLC-owned handshake step. SK: Dalsi neparny handshake krok vlastneny PLC.
   END_VAR
   NextState := NhExpectedState + 1;
   IF NhApiBuildNextFrame() THEN
      NhApiPublishFrame(NextState := NextState);
      NhApiPublishNextTargetFrame := TRUE;
   ELSE
      NhApiResetTransaction();
      NhApiPublishNextTargetFrame := FALSE;
   END_IF;
END_FUNCTION

FUNCTION NhApiPublishNextBroadcastFrame : BOOL
   // Publishes the next best-effort broadcast frame or returns to IDLE. SK: Publikuje dalsi best-effort broadcast ramec alebo sa vrati do IDLE.
   VAR
      NextState : UINT; // Next odd broadcast commit step. SK: Dalsi neparny broadcast commit krok.
   END_VAR
   IF NhExpectedState = 0 THEN
      NextState := 1;
   ELSE
      NextState := NhExpectedState + 2;
   END_IF;
   IF NhApiBuildNextFrame() THEN
      NhApiPublishFrame(NextState := NextState);
      NhApiPublishNextBroadcastFrame := TRUE;
   ELSE
      NhApiResetTransaction();
      NhApiPublishNextBroadcastFrame := FALSE;
   END_IF;
END_FUNCTION

FUNCTION NhApiProcessRx : BOOL
   // Validates the committed shared RX frame, executes it and publishes the first response frame. SK: Overi potvrdeny spolocny RX ramec, vykona ho a publikuje prvy ramec odpovede.
   VAR
      Buffer       : PTR_TO BYTE; // Byte view of NhApiRX. SK: Bajtovy pohlad na NhApiRX.
      TotalSize    : UINT;        // Declared complete RX size. SK: Deklarovana celkova velkost RX.
      PayloadSize  : UDINT;       // Declared payload size. SK: Deklarovana velkost payloadu.
      MessageType  : UINT;        // RX NH_API_MSG_* value. SK: RX hodnota NH_API_MSG_*.
      ExpectedCrc  : DWORD;       // CRC carried by RX header. SK: CRC ulozene v RX hlavicke.
      ActualCrc    : DWORD;       // CRC calculated by PLC. SK: CRC vypocitane PLC.
      ValidFrame   : BOOL;        // Header, size, owner and CRC are valid. SK: Hlavicka, velkost, vlastnik a CRC su platne.
      ConfigRecord : NH_ROOM_CONFIG; // Decoded config record. SK: Dekodovany config zaznam.
      StateRecord  : NH_ROOM_STATE;  // Decoded state record. SK: Dekodovany state zaznam.
      SourceRoomId : UDINT;       // Source ID of COPY_ROOM. SK: Zdrojove ID COPY_ROOM.
   END_VAR
   Buffer := ADR(NhApiRX);
   NhCommandResult := NH_API_RESULT_BAD_FRAME;
   ValidFrame := FALSE;
   TotalSize := UDINT_TO_UINT(NhApiReadU32(Buffer := Buffer, Offset := 28));
   PayloadSize := NhApiReadU32(Buffer := Buffer, Offset := 24);
   IF (TotalSize >= NH_API_HEADER_SIZE) AND (TotalSize <= NH_API_RX_BYTE_CAPACITY) AND
      (NhApiReadU32(Buffer := Buffer, Offset := 0) = DWORD_TO_UDINT(NH_API_MAGIC)) AND
      (NhApiReadU16(Buffer := Buffer, Offset := 4) = NH_API_VERSION) AND
      (NhApiReadU16(Buffer := Buffer, Offset := 6) = NH_API_HEADER_SIZE) AND
      (NhApiReadU32(Buffer := Buffer, Offset := 12) = NhActiveOwnerClientId) AND
      ((PayloadSize + UINT_TO_UDINT(NH_API_HEADER_SIZE)) = UINT_TO_UDINT(TotalSize)) THEN
      ExpectedCrc := UDINT_TO_DWORD(NhApiReadU32(Buffer := Buffer, Offset := 36));
      ActualCrc := NhApiFrameCrc32(Buffer := Buffer, Length := TotalSize);
      ValidFrame := ExpectedCrc = ActualCrc;
   END_IF;

   IF NOT ValidFrame THEN
      NhTransactionMode := NH_API_MODE_COMMAND;
      NhResultPending := TRUE;
      NhPendingConfigCount := 0;
      NhPendingStateCount := 0;
      NhApiPublishNextTargetFrame();
      NhApiProcessRx := FALSE;
      RETURN;
   END_IF;

   MessageType := NhApiReadU16(Buffer := Buffer, Offset := 8);
   CASE MessageType OF
      NH_API_MSG_SNAPSHOT_REQUEST:
         IF PayloadSize = 0 THEN
            NhCommandResult := NH_API_RESULT_OK;
            NhApiStartSnapshot();
            NhTransactionMode := NH_API_MODE_SNAPSHOT;
            NhApiPublishNextTargetFrame();
            NhApiProcessRx := TRUE;
            RETURN;
         END_IF;

      NH_API_MSG_ADD_ROOM:
         IF PayloadSize = UINT_TO_UDINT(NH_API_CONFIG_RECORD_SIZE) THEN
            NhApiReadConfigRecord(Buffer := Buffer, Offset := NH_API_HEADER_SIZE, Record := ConfigRecord);
            NhCommandResult := NhApiApplyAdd(Record := ConfigRecord);
         END_IF;

      NH_API_MSG_DELETE_ROOM:
         IF PayloadSize = 4 THEN
            NhCommandResult := NhApiApplyDelete(RoomId := NhApiReadU32(Buffer := Buffer, Offset := NH_API_HEADER_SIZE));
         END_IF;

      NH_API_MSG_COPY_ROOM:
         IF PayloadSize = (UINT_TO_UDINT(NH_API_CONFIG_RECORD_SIZE) + 4) THEN
            SourceRoomId := NhApiReadU32(Buffer := Buffer, Offset := NH_API_HEADER_SIZE);
            NhApiReadConfigRecord(Buffer := Buffer, Offset := NH_API_HEADER_SIZE + 4, Record := ConfigRecord);
            NhCommandResult := NhApiApplyCopy(SourceRoomId := SourceRoomId, Target := ConfigRecord);
         END_IF;

      NH_API_MSG_SET_ROOM_CONFIG:
         IF PayloadSize = UINT_TO_UDINT(NH_API_CONFIG_RECORD_SIZE) THEN
            NhApiReadConfigRecord(Buffer := Buffer, Offset := NH_API_HEADER_SIZE, Record := ConfigRecord);
            NhCommandResult := NhApiApplyConfig(Record := ConfigRecord);
         END_IF;

      NH_API_MSG_SET_ROOM_STATE:
         IF PayloadSize = UINT_TO_UDINT(NH_API_STATE_RECORD_SIZE) THEN
            NhApiReadStateRecord(Buffer := Buffer, Offset := NH_API_HEADER_SIZE, Record := StateRecord);
            NhCommandResult := NhApiApplyState(Record := StateRecord);
         END_IF;

      ELSE
         NhCommandResult := NH_API_RESULT_UNSUPPORTED;
   END_CASE;

   NhApiCaptureAllChanges();
   NhResultPending := TRUE;
   NhTransactionMode := NH_API_MODE_COMMAND;
   NhApiPublishNextTargetFrame();
   NhApiProcessRx := NhCommandResult = NH_API_RESULT_OK;
END_FUNCTION

FUNCTION NhApiProcessTest : BOOL
   // Applies one WebMaker/debug test action when the global API is free. SK: Vykona jednu WebMaker/debug testovaciu akciu, ked je globalne API volne.
   VAR
      Slot         : UINT;           // Located room slot. SK: Najdeny room slot.
      Index        : UINT;           // LOAD_800 model device index. SK: Index modeloveho zariadenia LOAD_800.
      StartMs      : UDINT;          // Scene application start time. SK: Cas zaciatku vykonania sceny.
      ConfigRecord : NH_ROOM_CONFIG; // Constructed config record. SK: Zostaveny config zaznam.
      StateRecord  : NH_ROOM_STATE;  // Constructed state record. SK: Zostaveny state zaznam.
   END_VAR
   NhApiProcessTest := FALSE;
   IF NOT NhApiTest.Execute THEN RETURN; END_IF;
   NhApiTest.Finished := FALSE;
   NhCommandResult := NH_API_RESULT_UNSUPPORTED;

   IF NhApiTest.Action = NH_API_TEST_REQUEST_SNAPSHOT THEN
      NhActiveOwnerClientId := 0;
      NhApiStartSnapshot();
      NhTransactionMode := NH_API_MODE_BROADCAST_SNAPSHOT;
      NhCommandResult := NH_API_RESULT_OK;
      NhApiPublishNextBroadcastFrame();
   ELSIF NhApiTest.Action = NH_API_TEST_AWAY THEN
      StartMs := NhApiSystemTimeMs();
      FOR Index := 1 TO 640 DO
         IF NhApiTest.Presence THEN
            IF Index <= 300 THEN
               NhLoadDevices[Index] := 16#01000000;
            ELSIF Index <= 420 THEN
               NhLoadDevices[Index] := 16#02000000;
            ELSIF Index <= 520 THEN
               NhLoadDevices[Index] := 16#030000AA;
            ELSIF Index <= 600 THEN
               NhLoadDevices[Index] := 16#040000B4;
            ELSE
               NhLoadDevices[Index] := 16#05000000;
            END_IF;
         ELSE
            IF Index <= 300 THEN
               NhLoadDevices[Index] := 16#01000064;
            ELSIF Index <= 420 THEN
               NhLoadDevices[Index] := 16#02000064;
            ELSIF Index <= 520 THEN
               NhLoadDevices[Index] := 16#030000D2;
            ELSIF Index <= 600 THEN
               NhLoadDevices[Index] := 16#040000DC;
            ELSE
               NhLoadDevices[Index] := 16#05000001;
            END_IF;
         END_IF;
      END_FOR;
      NhLoadTest.DepartureActive := NhApiTest.Presence;
      NhLoadTest.LastChangedCount := 640;
      NhLoadTest.LastApplyMs := NhApiSystemTimeMs() - StartMs;
      NhLoadTest.Sequence := NhLoadTest.Sequence + 1;
      NhCommandResult := NH_API_RESULT_OK;
   ELSIF NhApiTest.Action = NH_API_TEST_DELETE_ROOM THEN
      NhCommandResult := NhApiApplyDelete(RoomId := NhApiTest.RoomId);
   ELSIF NhApiTest.Action = NH_API_TEST_SET_STATE THEN
      Slot := NhApiFindRoom(RoomId := NhApiTest.RoomId);
      IF Slot = 0 THEN
         NhCommandResult := NH_API_RESULT_NOT_FOUND;
      ELSE
         StateRecord := NhRoomsState[Slot];
         StateRecord.Temperature := NhApiTest.Temperature;
         StateRecord.Humidity := NhApiTest.Humidity;
         StateRecord.Presence := NhApiTest.Presence;
         StateRecord.DayPhase := NhApiTest.DayPhase;
         StateRecord.CategoryMask := NhApiTest.CategoryMask;
         StateRecord.AlarmLevel := NhApiTest.AlarmLevel;
         StateRecord.Online := NhApiTest.Online;
         StateRecord.Twilight := NhApiTest.Twilight;
         NhCommandResult := NhApiApplyState(Record := StateRecord);
      END_IF;
   ELSE
      ConfigRecord.Used := TRUE;
      ConfigRecord.RoomId := NhApiTest.RoomId;
      ConfigRecord.Name := NhApiTest.Name;
      ConfigRecord.ProjectName := NhApiTest.ProjectName;
      ConfigRecord.IconId := NhApiTest.IconId;
      ConfigRecord.SortDefault := 0;
      IF NhApiTest.Action = NH_API_TEST_ADD_ROOM THEN
         NhCommandResult := NhApiApplyAdd(Record := ConfigRecord);
      ELSIF NhApiTest.Action = NH_API_TEST_COPY_ROOM THEN
         NhCommandResult := NhApiApplyCopy(SourceRoomId := NhApiTest.SourceRoomId, Target := ConfigRecord);
      ELSIF NhApiTest.Action = NH_API_TEST_SET_CONFIG THEN
         Slot := NhApiFindRoom(RoomId := NhApiTest.RoomId);
         IF Slot = 0 THEN
            NhCommandResult := NH_API_RESULT_NOT_FOUND;
         ELSE
            ConfigRecord.SortDefault := NhRoomsConfig[Slot].SortDefault;
            NhCommandResult := NhApiApplyConfig(Record := ConfigRecord);
         END_IF;
      END_IF;
   END_IF;

   IF (NhApiTest.Action <> NH_API_TEST_REQUEST_SNAPSHOT) AND NhApiCaptureAllChanges() THEN
      NhActiveOwnerClientId := 0;
      NhTransactionMode := NH_API_MODE_BROADCAST_DIFF;
      NhApiPublishNextBroadcastFrame();
   END_IF;
   NhApiTest.ResultCode := NhCommandResult;
   NhApiTest.Execute := FALSE;
   NhApiTest.Finished := TRUE;
   NhApiProcessTest := TRUE;
END_FUNCTION

FUNCTION NhApiCycle : BOOL
   // Executes one deterministic step of the global handshake every PLC cycle. SK: V kazdom PLC cykle vykona jeden deterministicky krok globalneho handshake.
   VAR
      NowMs      : UDINT; // Current PLC system time. SK: Aktualny systemovy cas PLC.
      ClientStep : UINT;  // State value written by the owner. SK: Hodnota State zapisana vlastnikom.
   END_VAR
   NowMs := NhApiSystemTimeMs();
   NhApiInfo.ApiVersion := NH_API_VERSION;

   // Internal ExpectedState is authoritative; a foreign write of State=0 may not abort an active transaction. SK: Interny ExpectedState je autorita; cudzi zapis State=0 nesmie prerusit aktivnu transakciu.
   IF NhExpectedState = NH_API_STATE_IDLE THEN
      NhExpectedState := NH_API_STATE_IDLE;
      NhActiveOwnerClientId := 0;
      NhApiInfo.State := NH_API_STATE_IDLE;
      IF NhApiInfo.OwnerClientId <> 0 THEN
         // The last OwnerClientId visible in this PLC cycle wins the claim. SK: Claim vyhra posledne OwnerClientId viditelne v tomto PLC cykle.
         NhActiveOwnerClientId := NhApiInfo.OwnerClientId;
         NhApiClearBuffer(Buffer := ADR(NhApiRX), Length := NH_API_RX_BYTE_CAPACITY);
         NhTransactionMode := NH_API_MODE_NONE;
         NhExpectedState := NH_API_STATE_OWNER_READY;
         NhTransactionLastMs := NowMs;
         NhApiInfo.State := NH_API_STATE_OWNER_READY;
         NhApiCycle := TRUE;
         RETURN;
      END_IF;

      IF NhApiTest.Execute THEN
         NhApiProcessTest();
         NhApiCycle := TRUE;
         RETURN;
      END_IF;

      IF NhApiCaptureAllChanges() THEN
         NhActiveOwnerClientId := 0;
         NhCommandResult := NH_API_RESULT_OK;
         NhTransactionMode := NH_API_MODE_BROADCAST_DIFF;
         NhApiPublishNextBroadcastFrame();
      END_IF;
      NhApiCycle := TRUE;
      RETURN;
   END_IF;

   IF NhActiveOwnerClientId <> 0 THEN
      IF (NowMs - NhTransactionLastMs) > NH_API_TRANSACTION_TIMEOUT_MS THEN
         NhApiResetTransaction();
         NhApiCycle := TRUE;
         RETURN;
      END_IF;

      // No other client may replace owner or State while this owner holds the transaction. SK: Ziadny iny klient nesmie pocas transakcie nahradit ownera ani State.
      IF NhApiInfo.OwnerClientId <> NhActiveOwnerClientId THEN
         NhApiInfo.OwnerClientId := NhActiveOwnerClientId;
         NhApiInfo.State := NhExpectedState;
         NhApiCycle := TRUE;
         RETURN;
      END_IF;

      IF NhApiInfo.State <> NhExpectedState THEN
         ClientStep := NhApiInfo.State;
         IF ClientStep = (NhExpectedState + 1) THEN
            NhExpectedState := ClientStep;
            NhTransactionLastMs := NowMs;
            IF ClientStep = NH_API_STATE_RX_READY THEN
               NhApiProcessRx();
            ELSIF (ClientStep MOD 2) = 0 THEN
               NhApiPublishNextTargetFrame();
            ELSE
               NhApiInfo.State := NhExpectedState;
            END_IF;
         ELSE
            NhApiInfo.State := NhExpectedState;
         END_IF;
      END_IF;
      NhApiCycle := TRUE;
      RETURN;
   END_IF;

   // OwnerClientId zero means a best-effort PLC broadcast with no per-client ACK. SK: Nulove OwnerClientId znamena best-effort PLC broadcast bez ACK jednotlivych klientov.
   NhApiInfo.OwnerClientId := 0;
   IF NhApiInfo.State <> NhExpectedState THEN NhApiInfo.State := NhExpectedState; END_IF;
   IF (NowMs - NhTransactionLastMs) >= NH_API_BROADCAST_HOLD_MS THEN
      NhApiPublishNextBroadcastFrame();
   END_IF;
   NhApiCycle := TRUE;
END_FUNCTION

(* ---- 04_Nh_Connect.st ---- *)
// NachHouse outbound transport pilot for CP-2000.
// The production protocol is binary NHAP; no PLCComS or TecoApi is used here.

VAR_GLOBAL
   NhConnectEnable        {PUBLIC_API} : BOOL := FALSE;
   NhConnectSendTest      {PUBLIC_API} : BOOL := FALSE;
   NhConnectConnected     {PUBLIC_API} : BOOL := FALSE;
   NhConnectReceived      {PUBLIC_API} : BOOL := FALSE;
   NhConnectError         {PUBLIC_API} : BOOL := FALSE;
   NhConnectRxLength      {PUBLIC_API} : UINT := 0;
   NhConnectSentBytes     {PUBLIC_API} : UDINT := 0;
   NhConnectReceivedBytes {PUBLIC_API} : UDINT := 0;
   NhConnectTestCounter   {PUBLIC_API} : UDINT := 0;
   NhConnectFrameCounter  {PUBLIC_API} : UDINT := 0;
   NhConnectCommandCounter {PUBLIC_API} : UDINT := 0;
   NhConnectRejectedCounter {PUBLIC_API} : UDINT := 0;
   NhConnectLastError     {PUBLIC_API} : STRING[80];
   NhConnectUrl           {PUBLIC_API} : STRING[255] := 'ws://192.168.33.113:18080/plc/load-800';
   NhConnectHeader        {PUBLIC_API} : STRING[80] := 'Authorization: Bearer local-test-token$0D$0A';
END_VAR

FUNCTION NhConnectCrc32 : DWORD
   VAR_INPUT
      Buffer : PTR_TO BYTE;
      Length : UINT;
   END_VAR
   VAR
      Crc : DWORD;
      Current : BYTE;
      Index : UINT;
      BitIndex : USINT;
   END_VAR
   Crc := 16#FFFFFFFF;
   IF Length > 0 THEN
      FOR Index := 0 TO Length - 1 DO
         Current := NhApiReadByte(Buffer := Buffer, Offset := Index);
         Crc := Crc XOR BYTE_TO_DWORD(Current);
         FOR BitIndex := 0 TO 7 DO
            IF (Crc AND 16#00000001) <> 0 THEN
               Crc := SHR(Crc, 1) XOR 16#EDB88320;
            ELSE
               Crc := SHR(Crc, 1);
            END_IF;
         END_FOR;
      END_FOR;
   END_IF;
   NhConnectCrc32 := NOT Crc;
END_FUNCTION

FUNCTION_BLOCK fbNhConnectPilot
   VAR_INPUT
      Enable : BOOL;
      SendTest : BOOL;
      ServerUrl : STRING[255];
      OptionalHeader : STRING[80];
   END_VAR
   VAR_OUTPUT
      Connected : BOOL;
      Received : BOOL;
      Error : BOOL;
      RxLength : UINT;
      SentBytes : UDINT;
      ReceivedBytes : UDINT;
      LastError : STRING[80];
   END_VAR
   VAR
      Socket : fbWebSocketClient;
      SendBuffer : ARRAY[1..MAX_LEN_WS_BUFFER] OF USINT;
      ReceiveBuffer : ARRAY[1..MAX_LEN_WS_BUFFER] OF USINT;
      SendEdge : R_TRIG;
      RequestSend : BOOL;
      ReceivePulse : BOOL;
      ReceiveLength : UINT;
      Index : UINT;
      LastPublishedFrameId : UDINT;
      FrameActive : BOOL;
      SendPhase : BOOL;
      FrameLength : UINT;
      FrameChecksum : DWORD;
      ChunkIndex : UINT;
      ChunkCount : UINT;
      ChunkOffset : UINT;
      ChunkLength : UINT;
      SourcePtr : PTR_TO BYTE;
      PendingCommand : ARRAY[0..255] OF BYTE;
      CommandPending : BOOL;
      CommandCommitted : BOOL;
      CommandLength : UINT;
      CommandOwner : UDINT;
      IncomingPayloadLength : UINT;
      IncomingChecksum : DWORD;
   END_VAR

   RequestSend := FALSE;
   SendEdge(CLK := SendTest);

   IF NOT Enable THEN
      FrameActive := FALSE;
      SendPhase := FALSE;
      LastPublishedFrameId := NhPublishedFrameId;
      CommandPending := FALSE;
      CommandCommitted := FALSE;
   END_IF;

   // Commit one received command through the existing V11 owner handshake.
   IF Enable AND CommandPending THEN
      IF NOT CommandCommitted AND (NhApiInfo.State = NH_API_STATE_OWNER_READY) AND
         (NhApiInfo.OwnerClientId = CommandOwner) THEN
         MemcpyPtr(Source := ADR(PendingCommand), Dest := ADR(NhApiRX), Length := UINT_TO_UDINT(CommandLength));
         NhApiInfo.State := NH_API_STATE_RX_READY;
         CommandCommitted := TRUE;
      ELSIF CommandCommitted AND (NhApiInfo.State = NH_API_STATE_IDLE) THEN
         CommandPending := FALSE;
         CommandCommitted := FALSE;
      END_IF;
   END_IF;

   // Capture every new V11 application frame and wrap it in NHAP Connect chunks.
   IF Enable AND Socket.isConnected AND NOT FrameActive AND
      (NhPublishedFrameId <> 0) AND (NhPublishedFrameId <> LastPublishedFrameId) THEN
      FrameLength := UDINT_TO_UINT(NhApiReadU32(Buffer := ADR(NhApiTX), Offset := 28));
      IF (FrameLength >= NH_API_HEADER_SIZE) AND (FrameLength <= NH_API_TX_BYTE_CAPACITY) THEN
         FrameChecksum := NhConnectCrc32(Buffer := ADR(NhApiTX), Length := FrameLength);
         ChunkCount := (FrameLength + 1407) / 1408;
         ChunkIndex := 0;
         FrameActive := TRUE;
         SendPhase := FALSE;
      ELSE
         LastPublishedFrameId := NhPublishedFrameId;
      END_IF;
   END_IF;

   IF Enable AND Socket.isConnected AND FrameActive AND NOT SendPhase THEN
      ChunkOffset := ChunkIndex * 1408;
      ChunkLength := FrameLength - ChunkOffset;
      IF ChunkLength > 1408 THEN ChunkLength := 1408; END_IF;

      NhApiWriteByte(Buffer := ADR(SendBuffer), Offset := 0, Value := 16#4E);
      NhApiWriteByte(Buffer := ADR(SendBuffer), Offset := 1, Value := 16#48);
      NhApiWriteByte(Buffer := ADR(SendBuffer), Offset := 2, Value := 16#41);
      NhApiWriteByte(Buffer := ADR(SendBuffer), Offset := 3, Value := 16#50);
      NhApiWriteByte(Buffer := ADR(SendBuffer), Offset := 4, Value := 1);
      NhApiWriteByte(Buffer := ADR(SendBuffer), Offset := 5, Value := 12); // V11 application frame
      NhApiWriteByte(Buffer := ADR(SendBuffer), Offset := 6, Value := BOOL_TO_BYTE(ChunkCount > 1));
      NhApiWriteByte(Buffer := ADR(SendBuffer), Offset := 7, Value := 32);
      NhApiWriteU32(Buffer := ADR(SendBuffer), Offset := 8, Value := NhPublishedFrameId);
      NhApiWriteU32(Buffer := ADR(SendBuffer), Offset := 12, Value := NhPublishedFrameId);
      NhApiWriteU16(Buffer := ADR(SendBuffer), Offset := 16, Value := ChunkIndex);
      NhApiWriteU16(Buffer := ADR(SendBuffer), Offset := 18, Value := ChunkCount);
      NhApiWriteU16(Buffer := ADR(SendBuffer), Offset := 20, Value := ChunkLength);
      NhApiWriteU16(Buffer := ADR(SendBuffer), Offset := 22, Value := 0);
      NhApiWriteU32(Buffer := ADR(SendBuffer), Offset := 24, Value := UINT_TO_UDINT(FrameLength));
      NhApiWriteU32(Buffer := ADR(SendBuffer), Offset := 28, Value := DWORD_TO_UDINT(FrameChecksum));
      SourcePtr := ADR(NhApiTX) + UINT_TO_UDINT(ChunkOffset);
      MemcpyPtr(Source := SourcePtr, Dest := ADR(SendBuffer[33]), Length := UINT_TO_UDINT(ChunkLength));
      RequestSend := TRUE;
      SendPhase := TRUE;
      NhConnectFrameCounter := NhConnectFrameCounter + 1;
   ELSIF FrameActive AND SendPhase THEN
      SendPhase := FALSE;
      ChunkIndex := ChunkIndex + 1;
      IF ChunkIndex >= ChunkCount THEN
         LastPublishedFrameId := NhPublishedFrameId;
         FrameActive := FALSE;
         // A targeted V11 response is acknowledged only after its last physical chunk was sent.
         IF (NhActiveOwnerClientId <> 0) AND ((NhApiInfo.State MOD 2) = 1) THEN
            NhApiInfo.State := NhApiInfo.State + 1;
         END_IF;
      END_IF;
   END_IF;

   IF Enable AND Socket.isConnected AND NOT FrameActive AND SendEdge.Q THEN
      // Minimal NHAP v1 HEARTBEAT frame. Header is 32 bytes, payload is empty.
      SendBuffer[1] := 16#4E; // N
      SendBuffer[2] := 16#48; // H
      SendBuffer[3] := 16#41; // A
      SendBuffer[4] := 16#50; // P
      SendBuffer[5] := 1;
      SendBuffer[6] := 30;
      SendBuffer[7] := 0;
      SendBuffer[8] := 32;
      NhConnectTestCounter := NhConnectTestCounter + 1;
      MemcpyPtr(Source := ADR(NhConnectTestCounter), Dest := ADR(SendBuffer[9]), Length := 4);
      FOR Index := 13 TO 32 DO
         SendBuffer[Index] := 0;
      END_FOR;
      SendBuffer[19] := 1;
      SendBuffer[20] := 0;
      RequestSend := TRUE;
   END_IF;

   Socket(
      rqConnect := Enable,
      serverUrl := ServerUrl,
      wsOptHeader := OptionalHeader,
      textMode := FALSE,
      pingTime := T#20s,
      rqSend := RequestSend,
      lenSend := SEL(FrameActive, 32, ChunkLength + 32),
      logSizeKB := 0,
      logMode := ONE_TIME_LOG,
      logFileName := 'NH_CONNECT.LOG',
      sendBuf := void(SendBuffer),
      recvBuf := void(ReceiveBuffer),
      isRecv => ReceivePulse,
      lenRecv => ReceiveLength
   );

   Connected := Socket.isConnected;
   Received := ReceivePulse;
   Error := Socket.isError;
   RxLength := ReceiveLength;
   SentBytes := Socket.sumaSend;
   ReceivedBytes := Socket.sumaRecv;
   LastError := Socket.lastErrDesc;

   // Commands are at most 256 bytes, therefore one physical WebSocket frame is sufficient.
   IF Enable AND ReceivePulse AND NOT CommandPending THEN
      IncomingPayloadLength := NhApiReadU16(Buffer := ADR(ReceiveBuffer), Offset := 20);
      IncomingChecksum := UDINT_TO_DWORD(NhApiReadU32(Buffer := ADR(ReceiveBuffer), Offset := 28));
      IF (ReceiveLength >= 72) AND
         (NhApiReadU32(Buffer := ADR(ReceiveBuffer), Offset := 0) = DWORD_TO_UDINT(NH_API_MAGIC)) AND
         (NhApiReadByte(Buffer := ADR(ReceiveBuffer), Offset := 4) = 1) AND
         (NhApiReadByte(Buffer := ADR(ReceiveBuffer), Offset := 5) = 20) AND
         (NhApiReadByte(Buffer := ADR(ReceiveBuffer), Offset := 7) = 32) AND
         (NhApiReadU16(Buffer := ADR(ReceiveBuffer), Offset := 16) = 0) AND
         (NhApiReadU16(Buffer := ADR(ReceiveBuffer), Offset := 18) = 1) AND
         (IncomingPayloadLength >= NH_API_HEADER_SIZE) AND
         (IncomingPayloadLength <= NH_API_RX_BYTE_CAPACITY) AND
         (ReceiveLength = IncomingPayloadLength + 32) AND
         (NhApiReadU32(Buffer := ADR(ReceiveBuffer), Offset := 24) = UINT_TO_UDINT(IncomingPayloadLength)) AND
         (NhConnectCrc32(Buffer := ADR(ReceiveBuffer[33]), Length := IncomingPayloadLength) = IncomingChecksum) THEN
         CommandOwner := NhApiReadU32(Buffer := ADR(ReceiveBuffer[33]), Offset := 12);
         IF (CommandOwner <> 0) AND (NhApiInfo.State = NH_API_STATE_IDLE) THEN
            CommandLength := IncomingPayloadLength;
            MemcpyPtr(Source := ADR(ReceiveBuffer[33]), Dest := ADR(PendingCommand), Length := UINT_TO_UDINT(CommandLength));
            CommandPending := TRUE;
            CommandCommitted := FALSE;
            NhApiInfo.OwnerClientId := CommandOwner;
            NhConnectCommandCounter := NhConnectCommandCounter + 1;
         ELSE
            NhConnectRejectedCounter := NhConnectRejectedCounter + 1;
         END_IF;
      ELSE
         NhConnectRejectedCounter := NhConnectRejectedCounter + 1;
      END_IF;
   END_IF;
END_FUNCTION_BLOCK

(* ---- prgMain.ST ---- *)
VAR_GLOBAL
   // Test PLC deployment only. Upload and verify this file before requesting activation.
   NhDeployRequest {PUBLIC_API} : BOOL := FALSE;
   NhDeployResult  {PUBLIC_API} : USINT := 0; // 0=none, 1=call returned TRUE, 2=API busy, 3=call returned FALSE (not final outcome)
   NhDeployBuild   {PUBLIC_API} : UDINT := 2026100251;
END_VAR

PROGRAM prgMain
   // Starts the API once and advances its handshake in every PLC cycle. SK: Jednorazovo spusti API a v kazdom PLC cykle posunie jeho handshake.
   VAR_INPUT
   END_VAR
   VAR_OUTPUT
   END_VAR
   VAR
      deployStarted : BOOL := FALSE;
      deployAccepted : BOOL;
      fileTransportOk : BOOL;
      jsonTestOk : BOOL;
      NhConnect : fbNhConnectPilot;
   END_VAR
   VAR_TEMP
   END_VAR

   NhApiInitialize();
   NhRxTextTransportCycle();
   NhApiCycle();
   fileTransportOk := NhFileTransportCycle();
   jsonTestOk := NhJsonTestCycle();

   NhConnect(
      Enable := NhConnectEnable,
      SendTest := NhConnectSendTest,
      ServerUrl := NhConnectUrl,
      OptionalHeader := NhConnectHeader,
      Connected => NhConnectConnected,
      Received => NhConnectReceived,
      Error => NhConnectError,
      RxLength => NhConnectRxLength,
      SentBytes => NhConnectSentBytes,
      ReceivedBytes => NhConnectReceivedBytes,
      LastError => NhConnectLastError
   );

   // Never deploy on the first cycle or repeat a request automatically.
   IF NOT deployStarted THEN
      NhDeployRequest := FALSE;
      NhDeployResult := 0;
      deployStarted := TRUE;
   ELSIF NhDeployRequest THEN
      NhDeployRequest := FALSE;
      IF NhApiInfo.State <> 0 THEN
         NhDeployResult := 2;
      ELSE
         deployAccepted := LoadNewPackage2(rq := TRUE, pckg := '//WWW/UPLOAD/NEW_PACK.TTR');
         IF deployAccepted THEN
            NhDeployResult := 1;
         ELSE
            NhDeployResult := 3;
         END_IF;
      END_IF;
   END_IF;
END_PROGRAM
